Fanuc KAREL source: kt00724.KL

PROGRAM KT00724
%STACKSIZE=65535
%PRIORITY=65535
%NOLOCKGROUP
VAR
P1 : JOINTPOS9
P2 : JOINTPOS9
OUT : BOOLEAN
BEGIN
-- UNRESOLVED_PC line 8 opcodes [22 63 23] marker_code=0
END KT00724
